(* IEC 61131-3 sources: HappyLearnCodesys/content/softmotion/CNC01_direct, 1 file *)

(* ---- Ipo.st ---- *)
PROGRAM Ipo
VAR
	trafo: SMC_TRAFO_Gantry2;
	p1,p2: SMC_ControlAxisByPos;
	trafof: SMC_TRAFOF_Gantry2;
	smci: SMC_Interpolator;
	mcp1, mcp2: MC_Power;
END_VAR
